// TIA Portal V17 export
// export: Created 2026-11-08T05:50:28.810374Z, ExportSetting WithDefaults, DisplayName Totally Integrated Automation Portal, DisplayVersion V17, DisplayName TIA Portal Openness, DisplayVersion V17, DisplayName TIA Portal Version Control Interface, DisplayVersion V17, DisplayName STEP 7 Professional, DisplayVersion V17, DisplayName STEP 7 Safety, DisplayVersion V17, DisplayName WinCC Professional, DisplayVersion V17
FUNCTION_BLOCK "FB_Motor_Moore"   // FB5, LAD
TITLE = Arranque y paro: máquina de estados MOORE
{ S7_Optimized_Access := 'TRUE' }
VERSION : 0.1
// Moore: las salidas dependen solo del estado. Generado por TIA_MCP_V17 (crear_maquina_estados).
// stored: AutoNumber true, IsIECCheckEnabled false, IsRetainMemResEnabled false, MemoryReserve 100, SetENOAutomatically false, UDAEnableTagReadback false
   VAR_INPUT
      Marcha : Bool;   // Orden de marcha (pulsador o HMI)
      Paro : Bool;   // Orden de paro: 1 = parar
      Termico_OK : Bool;   // 1 = relé térmico sin falla
      Reset : Bool;   // Reset de falla
   END_VAR
   VAR_OUTPUT
      Motor : Bool;   // Orden al contactor
      Piloto_Marcha : Bool;   // Piloto verde
      Piloto_Falla : Bool;   // Piloto rojo
      Estado : Int;   // Estado actual
   END_VAR
   VAR
      Estado_Actual : Int := 0;   // Estado de la máquina
   END_VAR
   VAR_TEMP
      Estado_Previo : Int;   // Estado al inicio del ciclo
   END_VAR
BEGIN

REGION Network 1: Foto del estado al inicio del ciclo
   // Las transiciones se evalúan sobre esta copia: un solo salto por ciclo.
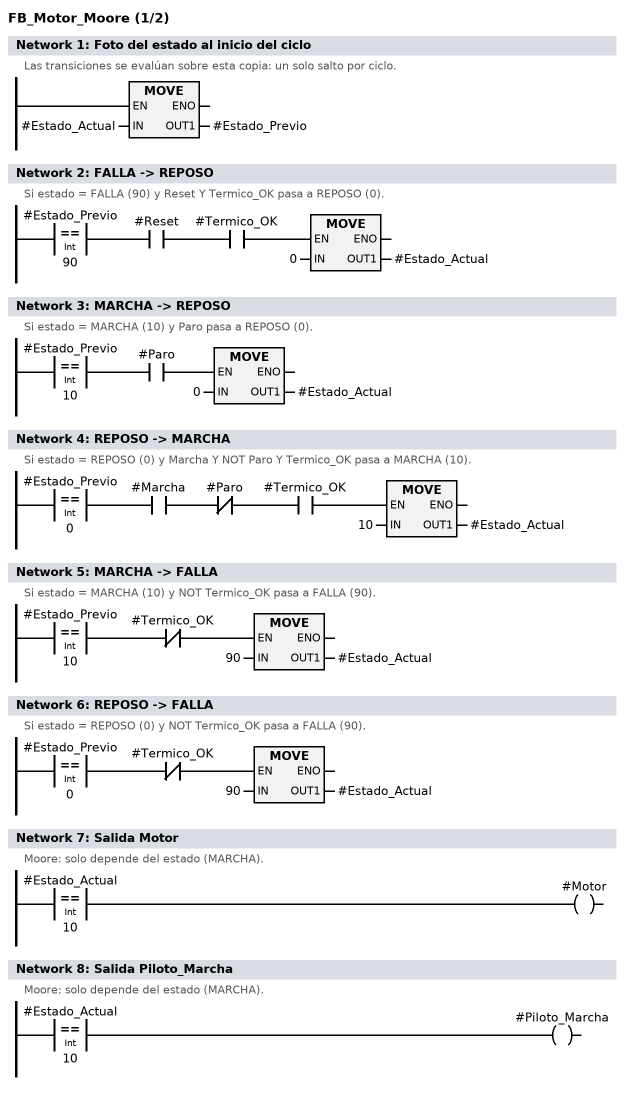
   RUNG wire#powerrail
      { S7_GenerateENO := "TRUE" } Move(in := #Estado_Actual, out1 => #Estado_Previo)
   END_RUNG
   // the same network as SCL:
   #Estado_Previo := #Estado_Actual;
END_REGION

REGION Network 2: FALLA -> REPOSO
   // Si estado = FALLA (90) y Reset Y Termico_OK pasa a REPOSO (0).
   RUNG wire#powerrail
      { S7_Templates := "SrcType := Int" } EQ_Contact(in1 := #Estado_Previo, in2 := 90)
      Contact( #Reset )
      Contact( #Termico_OK )
      { S7_GenerateENO := "TRUE" } Move(in := 0, out1 => #Estado_Actual)
   END_RUNG
   // the same network as SCL:
   IF (#Estado_Previo = 90) AND #Reset AND #Termico_OK THEN #Estado_Actual := 0; END_IF;
END_REGION

REGION Network 3: MARCHA -> REPOSO
   // Si estado = MARCHA (10) y Paro pasa a REPOSO (0).
   RUNG wire#powerrail
      { S7_Templates := "SrcType := Int" } EQ_Contact(in1 := #Estado_Previo, in2 := 10)
      Contact( #Paro )
      { S7_GenerateENO := "TRUE" } Move(in := 0, out1 => #Estado_Actual)
   END_RUNG
   // the same network as SCL:
   IF (#Estado_Previo = 10) AND #Paro THEN #Estado_Actual := 0; END_IF;
END_REGION

REGION Network 4: REPOSO -> MARCHA
   // Si estado = REPOSO (0) y Marcha Y NOT Paro Y Termico_OK pasa a MARCHA (10).
   RUNG wire#powerrail
      { S7_Templates := "SrcType := Int" } EQ_Contact(in1 := #Estado_Previo, in2 := 0)
      Contact( #Marcha )
      I_Contact( #Paro )
      Contact( #Termico_OK )
      { S7_GenerateENO := "TRUE" } Move(in := 10, out1 => #Estado_Actual)
   END_RUNG
   // the same network as SCL:
   IF (#Estado_Previo = 0) AND #Marcha AND NOT #Paro AND #Termico_OK THEN #Estado_Actual := 10; END_IF;
END_REGION

REGION Network 5: MARCHA -> FALLA
   // Si estado = MARCHA (10) y NOT Termico_OK pasa a FALLA (90).
   RUNG wire#powerrail
      { S7_Templates := "SrcType := Int" } EQ_Contact(in1 := #Estado_Previo, in2 := 10)
      I_Contact( #Termico_OK )
      { S7_GenerateENO := "TRUE" } Move(in := 90, out1 => #Estado_Actual)
   END_RUNG
   // the same network as SCL:
   IF (#Estado_Previo = 10) AND NOT #Termico_OK THEN #Estado_Actual := 90; END_IF;
END_REGION

REGION Network 6: REPOSO -> FALLA
   // Si estado = REPOSO (0) y NOT Termico_OK pasa a FALLA (90).
   RUNG wire#powerrail
      { S7_Templates := "SrcType := Int" } EQ_Contact(in1 := #Estado_Previo, in2 := 0)
      I_Contact( #Termico_OK )
      { S7_GenerateENO := "TRUE" } Move(in := 90, out1 => #Estado_Actual)
   END_RUNG
   // the same network as SCL:
   IF (#Estado_Previo = 0) AND NOT #Termico_OK THEN #Estado_Actual := 90; END_IF;
END_REGION

REGION Network 7: Salida Motor
   // Moore: solo depende del estado (MARCHA).
   RUNG wire#powerrail
      { S7_Templates := "SrcType := Int" } EQ_Contact(in1 := #Estado_Actual, in2 := 10)
      Coil( #Motor )
   END_RUNG
   // the same network as SCL:
   #Motor := #Estado_Actual = 10;
END_REGION

REGION Network 8: Salida Piloto_Marcha
   // Moore: solo depende del estado (MARCHA).
   RUNG wire#powerrail
      { S7_Templates := "SrcType := Int" } EQ_Contact(in1 := #Estado_Actual, in2 := 10)
      Coil( #Piloto_Marcha )
   END_RUNG
   // the same network as SCL:
   #Piloto_Marcha := #Estado_Actual = 10;
END_REGION

REGION Network 9: Salida Piloto_Falla
   // Moore: solo depende del estado (FALLA).
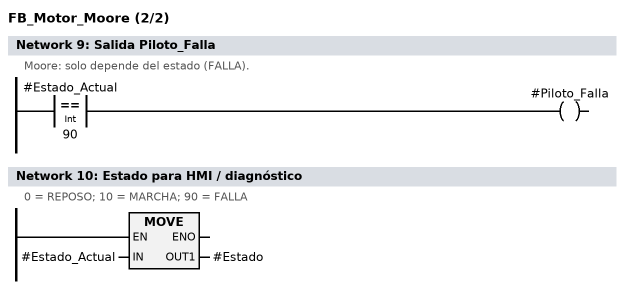
   RUNG wire#powerrail
      { S7_Templates := "SrcType := Int" } EQ_Contact(in1 := #Estado_Actual, in2 := 90)
      Coil( #Piloto_Falla )
   END_RUNG
   // the same network as SCL:
   #Piloto_Falla := #Estado_Actual = 90;
END_REGION

REGION Network 10: Estado para HMI / diagnóstico
   // 0 = REPOSO; 10 = MARCHA; 90 = FALLA
   RUNG wire#powerrail
      { S7_GenerateENO := "TRUE" } Move(in := #Estado_Actual, out1 => #Estado)
   END_RUNG
   // the same network as SCL:
   #Estado := #Estado_Actual;
END_REGION
END_FUNCTION_BLOCK
